  JIGs.append(create_jig_2(id=1, name="3FG", type=1, capacity=1, jig_offset=p[0,0,0,0,0,0]))
  JIGs.append(create_jig_2(id=2, name="jig input", type=2, capacity=1, jig_offset=p[0,0,0,0,0,-3.927]))
  JIGs.append(create_jig_2(id=3, name="jig output", type=3, capacity=1, jig_offset=p[0,0,0,0,0,0.78]))
  JIGs.append(create_jig_2(id=6, name="jig bin", type=6, capacity=1, jig_offset=p[0,0,0,0,0,0]))
  JIGs.append(create_jig_2(id=7, name="jig sarstedt racks", type=7, capacity=1, jig_offset=p[0,0,-0.02,0,0,0]))
  JIGs.append(create_jig_2(id=8, name="NoK Bin", type=8, capacity=1, jig_offset=p[0,0,0,0,0,0]))
  JIGs.append(create_jig_2(id=9, name="Pick bott jig", type=9, capacity=1, jig_offset=p[0,0,0,0,0,0]))
  JIGs.append(create_jig_2(id=10, name="Place bott jig", type=10, capacity=1, jig_offset=p[0,0,0,0,0,0]))
  JIGs.append(create_jig_2(id=11, name="bottle shake jig", type=11, capacity=1, jig_offset=p[0,0,0,0,0,0]))
  JIGs.append(create_jig_2(id=12, name="Pick Vial jig", type=12, capacity=1, jig_offset=p[0,0,0,0,0,0]))
  JIGs.append(create_jig_2(id=13, name="Place Vial jig", type=13, capacity=1, jig_offset=p[0,0,0,0,0,0]))
  JIGs.append(create_jig_2(id=14, name="Liquid transfer jig", type=14, capacity=1, jig_offset=p[0,0,0,0,0,0]))
  JIGs.append(create_jig_2(id=15, name="Pick station jig", type=15, capacity=1, jig_offset=p[0,0,0,0,0,0]))
  JIGs.append(create_jig_2(id=16, name="Place station jig", type=16, capacity=1, jig_offset=p[0,0,0,0,0,0]))
  JIGs.append(create_jig_2(id=17, name="Weigh station jig", type=17, capacity=1, jig_offset=p[0,0,0,0,0,0]))
  JIGs.append(create_jig_2(id=18, name="Pick station 1", type=18, capacity=1, jig_offset=p[0,0,0,0,0,0]))
  JIGs.append(create_jig_2(id=19, name="Pick station 2", type=19, capacity=1, jig_offset=p[0,0,0,0,0,0]))
  JIGs.append(create_jig_2(id=20, name="Pick station 3", type=20, capacity=1, jig_offset=p[0,0,0,0,0,0]))
  JIGs.append(create_jig_2(id=21, name="Tilt station jig", type=21, capacity=1, jig_offset=p[0,0,0,0,0,0]))
  $ 20 "Script: Powder_all_newspats.script"
  #global SERVER_IP   = "192.168.12.139"


  global tcp_dosing = p[0,0,0.15052,3.1415,0,0]
  global tcp_default = p[0,0,0.161,3.1415,0,0]

  global container_id = 0
  global powder_id  = 0
  global bulk_density = 0
  global H          = 0
  global H_c          = 0
  global mouth_d     = 0
  global mouth_sh    = 0
  global length_c     = 0
  global diameter   = 0
  global empty_weight_g  = 0
  global volume_ml    = 0
  global shape_code   = 0
  global flow_code   = 0
  global shape = ""
  global Flowability = ""
  global full_weight_g = 0
  global cent_edge = 0
  global pick_2_base = 0.2 # distance from tcp to base of picking table
  global wall_thickness = 0.002

  def read_db_data():

    socket_open(SERVER_IP, SERVER_PORT)
    sleep(0.5)
    socket_send_string("GET_DATACODE_FLOATS")
    sleep(5)

    local fl = socket_read_ascii_float(14)
    socket_close()

    global container_id = fl[1]
    global powder_id = fl[2]
    global bulk_density = fl[3]
    global H          = fl[4]/1000
    global H_c          = fl[5]/1000
    global mouth_d     = fl[6]/1000
    global mouth_sh    = fl[7]/1000
    global length_c     = fl[8]/1000
    global diameter   = fl[9]/1000
    global empty_weight_g = fl[10]
    global volume_ml    = fl[11]
    global full_weight_g = fl[12]
    global flow_code   = fl[13]
    global shape_code   = fl[14]

  	if (flow_code == 1.0):
  		global Flowability = "MEDIUM"
  	elif (flow_code == 2.0):
  		global Flowability = "LOW"
  	else:
  		global Flowability = "HIGH"
  	end

  	if ( shape_code == 1.0):
  		shape = "cylindrical"
  		cent_edge =  diameter
  	else:
  		shape = "cubical"
  		cent_edge =  length_c
  	end

  	read_spatula_data()

  end

  def send_picking_info(Pow_name, target_weight):
    socket_open(SERVER_IP, SERVER_PORT)
    cmd = "PICK:"+Pow_name+";"+to_str(target_weight)
    socket_send_string(cmd)
    sleep(0.1)
    socket_close()
  end

  #### POTS ####
  def tilt_send(angle):
  	socket_open(SERVER_IP, SERVER_PORT)
  	angle = 92.0 - angle
  	socket_send_string("TILT:"+to_str(angle))
  	sync()
  	sleep(0.5)
  	socket_close()
  end

  def CW_Rotate(angle):
  	socket_open(SERVER_IP, SERVER_PORT)
  	socket_send_string("CWROTATE:"+to_str(angle))
  	sync()
  	sleep(0.5)
  	socket_close()
  end

  def CCW_Rotate(angle):
  	socket_open(SERVER_IP, SERVER_PORT)
  	socket_send_string("CCWROTATE:"+to_str(angle))
  	sync()
  	sleep(0.5)
  	socket_close()
  end

  def CW_full_Rotate():
  	socket_open(SERVER_IP, SERVER_PORT)
  	socket_send_string("FULLROTATE:"+to_str(1))
  	sync()
  	sleep(0.5)
  	socket_close()
  end

  def CCW_full_Rotate():
  	socket_open(SERVER_IP, SERVER_PORT)
  	socket_send_string("FULLROTATE:"+to_str(-1))
  	sync()
  	sleep(0.5)
  	socket_close()
  end

  def tilt_to_home():
  	socket_open(SERVER_IP, SERVER_PORT)
  	socket_send_string("HOME")
  	sync()
  	sleep(0.5)
  	socket_close()
  end
  #######
  def vibration_1():
  	set_analog_out(0,0.4)
  	sleep(1)
  	set_analog_out(0,0.0)
  	sleep(0)
  end

  def vibration_2():
  	set_analog_out(0,0.4)
  	sleep(0.8)
  	set_analog_out(0,0.0)
  	sleep(0.2)
  end

  def vibration_3():
  	set_analog_out(0,0.4)
  	sleep(0.5)
  	set_analog_out(0,0.0)
  	sleep(0.3)
  end

  def vibration_4():
  	set_analog_out(0,0.4)
  	sleep(0.5)
  	set_analog_out(0, 0.0)
  	sleep(0.5)
  end

  def vibration_5():
  	set_analog_out(0,0.4)
  	sleep(0.2)
  	set_analog_out(0, 0.0)
  	sleep(0.8)
  end

  ##################

  global gear_2_holder = 0.018
  global hinge_2_base = 0.0421
  global TCP_2_tip_x = 0.0047
  global spatula_len = 0.182
  global spatula_offset = p[TCP_2_tip_x,0,spatula_len,0,0,0]
  global SPATULA_L_VOL_ML = 0.0
  global SPATULA_M_VOL_ML = 0.0
  global SPATULA_S_VOL_ML = 0.0
  global SPATULA_FLAT_M_VOL_ML  = 0.0
  global SPATULA_FLAT_S_VOL_ML  = 0.0

  global DB_SPATULA_L_DEPTH = 0.0
  global DB_SPATULA_M_DEPTH = 0.0
  global DB_SPATULA_S_DEPTH = 0.0
  global DB_SPATULA_FLAT_M_DEPTH = 0.0
  global DB_SPATULA_FLAT_S_DEPTH = 0.0
  global DB_SPATULA_L_MID = 0.0
  global DB_SPATULA_M_MID = 0.0
  global DB_SPATULA_S_MID = 0.0
  global DB_SPATULA_FLAT_M_MID = 0.0
  global DB_SPATULA_FLAT_S_MID = 0.0
  global DB_SPATULA_L_RY = 0.0
  global DB_SPATULA_M_RY = 0.0
  global DB_SPATULA_S_RY = 0.0
  global DB_SPATULA_FLAT_M_RY = 0.0
  global DB_SPATULA_FLAT_S_RY = 0.0

  def read_spatula_data():
  	socket_open(SERVER_IP, SERVER_PORT)
  	sleep(0.2)
  	socket_send_string("GET_SPATULA_FLOATS")
  	sleep(0.5)
  	local fl = socket_read_ascii_float(25)
  	socket_close()

  	global DB_SPATULA_L_DEPTH = fl[1]/1000
  	global DB_SPATULA_L_MID = fl[2]/2000
  	global SPATULA_L_VOL_ML = fl[3]
  	global DB_SPATULA_L_RY = fl[4]
  	global DB_SPATULA_M_DEPTH = fl[6]/1000
  	global DB_SPATULA_M_MID = fl[7]/2000
  	global SPATULA_M_VOL_ML = fl[8]
  	global DB_SPATULA_M_RY = fl[9]
  	global DB_SPATULA_S_DEPTH = fl[11]/1000
  	global DB_SPATULA_S_MID = fl[12]/2000
  	global SPATULA_S_VOL_ML = fl[13]
  	global DB_SPATULA_S_RY = fl[14]
  	global DB_SPATULA_FLAT_M_DEPTH = fl[16]/1000
  	global DB_SPATULA_FLAT_M_MID = fl[17]/2000
  	global SPATULA_FLAT_M_VOL_ML = fl[18]
  	global DB_SPATULA_FLAT_M_RY = fl[19]
  	global DB_SPATULA_FLAT_S_DEPTH = fl[21]/1000
  	global DB_SPATULA_FLAT_S_MID = fl[22]/2000
  	global SPATULA_FLAT_S_VOL_ML = fl[23]
  	global DB_SPATULA_FLAT_S_RY = fl[24]
  end

  def correction_reset():
  	global g_k = 0.0
  	global g_depth_corr = 0.0
  	global g_prev_cum_w = weight_value
  end

  def params_init():

  	global scoop_status= ""
  	global w_dosed_total = 0.0
  	global last_scale = 0.0
  	global tilt_angle_sent = 0.0
  	global level = 0.0
  	global target_g = 0.0
  	global angle_max = 65
  	global angle_min = 30
  	global gain_per_percent = (angle_max - angle_min)/100
  	global ry_deg_safe = 0
  	global ry_deg = 0
  	global delta_count=0

  	global scoop_ct = 0
  	global error_sum = 0.0
  	global error_sq_sum = 0.0
  	global scoop_g = 0.0

  	global g_k =0.0
  	global g_eta = 0.3

  	global g_gain_scale = 0.07
  	global g_k_min = 0.0
  	global g_k_max = 0.09

  	# ---------- Damping ----------
  	global g_alpha_under = 0.75   # aggressive when undershooting
  	global g_alpha_over  = 0.60   # conservative when overshooting

  	# ---------- Search ----------
  	global g_engagement_min = 0.05
  	global g_search_step = 0.01      # 3 mm

  	# ---------- Deadband ----------
  	global g_tol = 0.02               # 20 mg minimum
  	global g_tol_ratio = 0.05         # ±5% of target

  	# ---------- Limits ----------
  	global g_corr_max = 0.020         # 20 mm maximum correction

  	# ---------- States ----------
  	global g_depth_corr = 0.0
  	global g_prev_cum_w = -1.0
  	global z_ratio = 0.0
  	global z_offset = 0.0
  end

  def clamp(x, lo, hi):
  	if(x<lo):
  		return lo
  	elif (x>hi):
  		return hi
  	else:
  		return x
  	end
  end

  def compute_level_percent(W_now, weight_value):   # W_now = container+powder, weight_value = live scale reading
      global delta = weight_value - last_scale

      if (delta < 0.0):
          delta = 0.0
      end

      global w_dosed_total = w_dosed_total + delta
      global last_scale = weight_value     # update the last scale reading

      local W_eff = W_now - w_dosed_total
      if (W_eff <  empty_weight_g):
          W_eff =  empty_weight_g
      end

      # Compute powder level %
      level = 100.0 * (W_eff -  empty_weight_g) / (full_weight_g -  empty_weight_g)

      # Clamp to 0–100
      level = clamp(level, 0, 100)
    textmsg("deb 1 = ", level)
      return level
  end

  def deg2rad(d):
  	return d*3.141592/180
  end

  def my_abs(val):
  	if (val<0):
  		return -val
  	else:
  		return val
  	end
  end

  def compute_tilt_deg(level_percent):
  	angle = angle_min + gain_per_percent*(100.0-level_percent)

    	textmsg("deb 2 = ", angle)
  	return clamp(angle, angle_min, angle_max)
  end

  def tilt(level_percentage):
  	new_angle = compute_tilt_deg(level_percentage)
    	textmsg("deb angle 1 = ", new_angle)
  	global angle_rel = new_angle - tilt_angle_sent
    	textmsg("deb 2 = ", angle_rel)

  	if my_abs(angle_rel)>2.0:
    		textmsg("deb loop")
  		tilt_send(new_angle)
  		global angle_deg = new_angle
    		textmsg("deb 2 = ", angle_deg)
  		global tilt_angle_sent = new_angle
  		global p_center_vertical = center_pose()
  		global p_center = updated_center_pose(p_center_vertical, angle_deg)
  	end
    	textmsg("deb loop exit")

  	tilt_send(angle_deg)
    	textmsg("deb angle 2 =", angle_deg)

  end

  def compute_scoop_depth(level, weight_value, target_g):

      global scoop_depth_rel = ((100.0-level)/100.0)*(H-mouth_sh)

      if (g_prev_cum_w < 0):
          g_prev_cum_w = weight_value
          g_depth_corr = 0.0

      else:
          global scoop_g = weight_value - g_prev_cum_w
          g_prev_cum_w = weight_value

          local error = target_g - scoop_g
          local engagement = scoop_g / target_g

          local tol = g_tol_ratio * target_g
          if (tol < g_tol):
              tol = g_tol
          end
          if ((engagement < g_engagement_min) and (scoop_g < target_g)):
              g_depth_corr = g_depth_corr + g_search_step
          elif (my_abs(error) <= tol):
  			sync()
          else:
              local error_norm = my_abs(error / target_g)
              local g_target = clamp(g_gain_scale * error_norm,g_k_min,g_k_max)

              g_k = (1.0-g_eta) * g_k + g_eta * g_target
              if (error > 0):
                  local corr = g_k * error
                  g_depth_corr = g_depth_corr +g_alpha_under * corr
              else:
                  local corr = g_k * error
                  g_depth_corr = g_depth_corr +g_alpha_over * corr

              end
              g_depth_corr = clamp(g_depth_corr,-g_corr_max,g_corr_max)

          end
      end
      scoop_depth = scoop_depth_rel + g_depth_corr
      scoop_depth = clamp(scoop_depth, 0.0, H)
      return scoop_depth

  end

  def get_scoop_weight(spatula, bulk_density):

  	local vol = 0

  	if (spatula == "spatula_L"):
  		vol = SPATULA_L_VOL_ML
  		global spatula_depth = DB_SPATULA_L_DEPTH
  		global spatula_mid   = DB_SPATULA_L_MID
  		global spatula_ry    = DB_SPATULA_L_RY

  	elif (spatula == "spatula_M"):
  		vol = SPATULA_M_VOL_ML
  		global spatula_depth = DB_SPATULA_M_DEPTH
  		global spatula_mid   = DB_SPATULA_M_MID
  		global spatula_ry    = DB_SPATULA_M_RY

  	elif (spatula == "spatula_S"):
  		vol = SPATULA_S_VOL_ML
  		global spatula_depth = DB_SPATULA_S_DEPTH
  		global spatula_mid   = DB_SPATULA_S_MID
  		global spatula_ry    = DB_SPATULA_S_RY

  	elif (spatula == "spatula_flat_M"):
  		vol = SPATULA_FLAT_M_VOL_ML
  		global spatula_depth = DB_SPATULA_FLAT_M_DEPTH
  		global spatula_mid   = DB_SPATULA_FLAT_M_MID
  		global spatula_ry    = DB_SPATULA_FLAT_M_RY

  	elif (spatula == "spatula_flat_S"):
  		vol = SPATULA_FLAT_S_VOL_ML
  		global spatula_depth = DB_SPATULA_FLAT_S_DEPTH
  		global spatula_mid   = DB_SPATULA_FLAT_S_MID
  		global spatula_ry    = DB_SPATULA_FLAT_S_RY
  	else:
  		textmsg("Unknown spatula type")
  		return 0.0
  	end
  	global target_g = vol * bulk_density
  	return target_g

  end

  def select_spatula(Flowability, level, diff, bulk_density, mouth_d ):

      local k = 1.1
      global powder_height = (H  - mouth_sh ) * level/100

      if (Flowability == "LOW"):
          local gFM = get_scoop_weight("spatula_flat_M", bulk_density)
  		local mouth_ok_FM = (mouth_d >= 0.05)
  		local level_ok_FM = (spatula_mid  < powder_height)
          local diff_ok_FM  = (diff > k * gFM)
  		local flatM_ok = mouth_ok_FM and level_ok_FM and diff_ok_FM
          if (flatM_ok):
              return "spatula_flat_M"
          else:
              return "spatula_flat_S"
          end
      end

      local gL = get_scoop_weight("spatula_L", bulk_density)
      local mouth_ok_L = (mouth_d  >= 0.05)
      local level_ok_L = (spatula_mid < powder_height)
      local diff_ok_L  = (diff > k * gL)

      local large_ok = mouth_ok_L and level_ok_L and diff_ok_L
      local gM = get_scoop_weight("spatula_M", bulk_density)
      local level_ok_M = (spatula_mid < powder_height)
      local diff_ok_M  = (diff > k * gM)

      local medium_ok = level_ok_M and diff_ok_M

      if (large_ok):
          return "spatula_L"
      elif (medium_ok):
          return "spatula_M"
      else:
          return "spatula_S"
      end
  end

  def after_scoop():
  	set_tcp(tcp_dosing)
  	set_analog_out(0,0.0)
  	tilt_send(angle_deg)
  	sleep(0.5)
  	movel(lifted_pose, a=0.05, v=0.2)
  	movel(move_inside_spill, a=0.05, v=0.2)
  	set_analog_out(0,0.4)
  	if (Flowability == "LOW"):
  		movel(end_rel_tilted_level2, a=0.03, v=0.1)
  		sleep(0.5)
  		movel(move_inside_spill, a=0.05, v=0.2)
  	  	movel(pose_trans(move_inside_spill, p[0,0,0,0,0,2.0]), a=0.05, v=0.2)
  		#movel(tilted_pose_in_base2, a=0.05, v=0.2)
  	else:
  	    movel(pose_trans(move_inside_spill, p[0,0,0,0,0,2.0]), a=0.05, v=0.2)
  	    movel(move_inside_spill, a=0.05, v=0.2)
  	end
  	set_analog_out(0,0.0)
  	movel(lifted_pose, a=0.5, v=0.5)
  	tilt_to_home()
  	set_tcp(tcp_default)
  end

  def center_pose():
  	global p_translated = container_place
  	#global p_translated = pots_axis_temp

  	#cx = p_translated[0]
  	#cy = p_translated[1]
  	#cz = p_translated[2]

  	global p_center_vertical_temp = pose_trans(p_translated, p[0,0,0, deg2rad(90), 0, 0])
  	cx = p_center_vertical_temp[0]
  	cy = p_center_vertical_temp[1]
  	cz = p_center_vertical_temp[2]
  	rx = p_center_vertical_temp[3]
  	ry = p_center_vertical_temp[4]
  	rz = p_center_vertical_temp[5]

  	global p_center_vertical_temp = p[cx,cy,cz, 0, 0, rz]
  	trans_rel = p[0,0,-pick_2_base+H,0,0,0]
  	global p_center_vertical =  pose_trans(p_center_vertical_temp, trans_rel)
  	return p_center_vertical
  end

  def updated_center_pose(p_center_vertical, angle_deg):
  	hinge_pose = pose_trans(p_center_vertical, p[0,0,-hinge_2_base-gear_2_holder-H ,0,0,0])
  	local_rel = pose_trans(pose_inv(hinge_pose), p_center_vertical)

  	rot_tilt = p[0,0,0, -deg2rad(angle_deg),0,0]
  	local_rel_tilted = pose_trans(rot_tilt, local_rel)

  	global p_center = pose_trans(hinge_pose, local_rel_tilted)
  	return p_center
  end

  def scoop_powder(p_center):
  	vibration_voltage = 0.4
  	global scoop_radius_default = 0.0

  	scoop_radius_default = mouth_d /2 - spatula_depth - wall_thickness
  	scoop_safe_entry_pose = pose_trans(p_center, p[-TCP_2_tip_x,0,spatula_len+0.05,0,0,0])
  	scoop_entry_pose = pose_trans(p_center, p[-TCP_2_tip_x,0,spatula_len,0,0,0])

  	movel(scoop_safe_entry_pose, a=0.1, v=0.25)
  	movel(scoop_entry_pose, a=0.1, v=0.25)

  	scoop_start_rel_int = p[0, 0, -mouth_sh , 0, 0, 0]
  	scoop_start_pose_int = pose_trans(scoop_entry_pose, scoop_start_rel_int)


  	#local ry_deg = map_tilt_to_ry_deg(angle_deg,level)
  	#local ry_result = map_tilt_to_ry_deg(angle_deg,level)

  	#global scoop_depth = compute_scoop_depth(level,weight_value, target_g)

  	global ry = deg2rad(90-angle_deg)

  	#global ry_safe = ry_result[0]
  	#global ry = deg2rad(ry_result[1])

  	if (spatula_mid < powder_height):

  		global total_depth = mouth_sh + scoop_depth + spatula_mid
  		global total_depth = clamp(total_depth, 0, H - spatula_mid)

  		safe_scoop_pivot = (mouth_d  - spatula_depth-wall_thickness)/(total_depth)
  		global ry_safe = asin(safe_scoop_pivot)

  		scoop_start_rel = p[scoop_radius_default, 0, -total_depth, 0, 0, 0]

  		rot_mid = p[0, 0, 0, 0, 0, 0.785]
  		rot_end = p[0, 0, 0, 0, 0, 1.5708]

  		scoop_via_rel = pose_trans(rot_mid, scoop_start_rel)
  		scoop_end_rel = pose_trans(rot_end, scoop_start_rel)

  		scoop_start_pose = pose_trans(scoop_entry_pose, scoop_start_rel)
  		scoop_via_pose = pose_trans(scoop_entry_pose, scoop_via_rel)
  		scoop_end_pose = pose_trans(scoop_entry_pose, scoop_end_rel)


  			if (Flowability == "LOW" and level <= 50):
  				movel(pose_trans(scoop_start_pose_int,p[0,0,0,0,0,-1.5708]), a=0.1, v=0.25)
  				local spatula_base = pose_trans(scoop_entry_pose, p[0, 0, -H+wall_thickness, 0, 0, 0])
  				local scrape_pivot = pose_trans(scoop_entry_pose, p[0,0, -spatula_len,0,0,0])

  				global sticky_in_angle = -atan((cent_edge/2-spatula_depth)/H)
  				spatula_tilt_rel = pose_trans(pose_inv(scrape_pivot), spatula_base)

  				spatula_tilt = pose_trans(spatula_tilt_rel, p[0, 0, 0, 0, sticky_in_angle, 0])
  				global tilted_pose = pose_trans(scrape_pivot, p[0,0,0,spatula_tilt[3],spatula_tilt[4], spatula_tilt[5]])

  				global tilted_pose = pose_trans(tilted_pose, p[0,0,spatula_len-H+wall_thickness,0,0,0])
  				global rotate_90=pose_trans(tilted_pose,p[0,0,0,0,0,-1.5708])
  				movel(rotate_90,a=0.1, v=0.25)
  				CW_full_Rotate()
  				movel(scoop_start_pose, a=0.1, v=0.25)
  			else:
  				movel(scoop_start_pose_int, a=0.1, v=0.25)
  				movel(scoop_start_pose, a=0.1, v=0.25)
  				CW_full_Rotate()
  			end

  		movec(scoop_via_pose, scoop_end_pose, a=0.05, v=0.04)
  		#sleep(1.0)

  		# safe_retention
  		local pivot_pose = pose_trans(scoop_end_pose, p[0,0,total_depth-spatula_len,0,0,0])
  		local end_rel = pose_trans(pose_inv(pivot_pose), scoop_end_pose)
  		local end_rel_tilted = pose_trans(end_rel, p[0, 0, 0, 0, ry_safe-deg2rad(spatula_ry), 0])
  		local tilted_pose_in_base = pose_trans(pivot_pose, p[0,0,0,end_rel_tilted[3],end_rel_tilted[4], end_rel_tilted[5]])
  		local tilted_pose_in_base = pose_trans(tilted_pose_in_base, p[0, 0, spatula_len-total_depth, 0, 0, 0])
  		# sptula pivoted around the container rim of the mouth at ry_safe
  		movel(tilted_pose_in_base, a=0.03, v=0.1)

  		global safe_x = sin(ry_safe)*(total_depth-mouth_sh - (mouth_d - spatula_depth)*tan(ry_safe/2))
  		global safe_z = cos(ry_safe)*(total_depth-mouth_sh - (mouth_d - spatula_depth)*tan(ry_safe/2))

  		local safe_up = pose_trans(tilted_pose_in_base, p[-safe_x,0,safe_z,0,0,0])
  		movel(safe_up, a=0.03, v=0.1)

  		# full exit
  		local pivot_pose2 = pose_trans(scoop_entry_pose, p[0,0,-spatula_len,0,0,0])
  		local end_rel2 = pose_trans(pose_inv(pivot_pose2), tilted_pose_in_base)
  		#popup("is the spatula crashing front? ", blocking = True)
  		local end_rel_tilted2 = pose_trans(end_rel2, p[0, 0, 0, 0, ry-ry_safe-deg2rad(spatula_ry), 0])

  	else : # emptying logic
  		#CCW_full_Rotate()

  		spatula_base = pose_trans(scoop_entry_pose, p[0, 0, -H+wall_thickness, 0, 0, 0])
  		local pivot_pose2 = pose_trans(scoop_entry_pose, p[0,0,-spatula_len,0,0,0])
  		# tilt inwards
  		global in_angle = -atan((cent_edge/2-spatula_depth)/H)
  		spatula_tilt_rel = pose_trans(pose_inv(pivot_pose2), spatula_base)

  		spatula_tilt = pose_trans(spatula_tilt_rel, p[0, 0, 0, -in_angle, 0, 0])
  		global tilted_pose = pose_trans(pivot_pose2, p[0,0,0,spatula_tilt[3],spatula_tilt[4], spatula_tilt[5]])

  		global tilted_pose = pose_trans(tilted_pose, p[0,0,spatula_len-H+wall_thickness,0,0,0])

  		movel(tilted_pose,a=0.1, v=0.25)
  		CW_full_Rotate()
  		sleep(1)
  		rotate90=pose_trans(tilted_pose,p[0,0,0,0,0,1.5708])

  		#sleep(1)
  		#Rotate()
  		#sleep(0.2)
  		movel(rotate90, a=0.1, v=0.1)
  		#popup("is the spatula crashing front? ", blocking = True)
  		movel(pose_trans(scoop_start_pose_int,p[0,0,0,0,0,1.5708]), a=0.03, v=0.1)
  		# full exit
  		#local pivot_pose2 = pose_trans(scoop_entry_pose, p[0,0,-spatula_len,0,0,0])
  		local end_rel2 = pose_trans(pose_inv(scoop_entry_pose), rotate90)
  		local end_rel_tilted2 = pose_trans(end_rel2, p[0, 0, 0, 0, ry-in_angle-deg2rad(spatula_ry), 0])
  	end

  	# exit flat spoon
  	global tilted_pose_in_base2 = pose_trans(pivot_pose2, p[0,0,0,end_rel_tilted2[3],end_rel_tilted2[4], end_rel_tilted2[5]])
  	global tilted_pose_in_base2 = pose_trans(tilted_pose_in_base2, p[0, 0, spatula_len-spatula_mid, 0, 0, 0])
  	# spaula exited at center of the mouth at ry
  	movel(tilted_pose_in_base2, a=0.03, v=0.1)

  	if(spatula == "spatula_S"):
  		if(level>=80):
  			global z_ratio = 0.0
  		elif(level == 0.0):
  			global z_ratio = 1.0
  		else:
  			global z_ratio = (80-level)/80
  		end
  		z_offset = 4*spatula_mid*z_ratio
  	elif(spatula == "spatula_flat_S"):
  		if(level>=50):
  			global z_ratio = 0.0
  		elif(level == 0.0):
  			global z_ratio = 1.0
  		else:
  			global z_ratio = (50-level)/50
  		end
  		z_offset = 4*spatula_mid*z_ratio
  	else:
  	    z_offset = 0.0
  	end

  	global move_inside_spill = pose_trans(tilted_pose_in_base2, p[0,0,-z_offset,0,0,0])
  	movel(move_inside_spill, a=0.03, v=0.1)

  	if(scoop_status== "normal"):
  		vib_thread=True
  		if (spatula=="spatula_S"):
  			vibration_3()
  			local ry_level = deg2rad(5)
  		elif(spatula=="spatula_flat_S" or spatula=="spatula_flat_M"):
  			vibration_3()
  			local ry_level = deg2rad(5)
  		else:
  			set_analog_out(0,0.4)
  			local ry_level = deg2rad(15)
  		end

  		# remove excess
  		local pivot_pose_level = pose_trans(move_inside_spill, p[0,0,-spatula_len,0,0,0])
  		local end_rel_level = pose_trans(pose_inv(pivot_pose_level), move_inside_spill)
  		local end_rel_tilted_level = pose_trans(end_rel_level, p[0, 0, 0, 0, -ry_level, 0])
  		global end_rel_tilted_level2 = pose_trans(pivot_pose_level, p[0, 0, 0,end_rel_tilted_level[3],end_rel_tilted_level[4], end_rel_tilted_level[5]])
  		global end_rel_tilted_level2 = pose_trans(end_rel_tilted_level2, p[0,0,spatula_len,0,0,0])
  		movel(end_rel_tilted_level2, a=0.03, v=0.1)

  		if (spatula == "spatula_flat_S" or spatula == "spatula_flat_M"):
  			vib_thread=False
  			set_analog_out(0, 0.0)
  		end
  	else:
  		set_analog_out(0, 0.0)
  	end
  	movel(tilted_pose_in_base2, a=0.03, v=0.1)
  	set_analog_out(0, 0.0)
  	vib_thread=False
  	global lifted_pose = pose_trans(tilted_pose_in_base2, p[-0.04,0,0.04,0,0,0]) # safety distance away from the container

  	movel(lifted_pose, a=0.03, v=0.1)
  	tilt_to_home()
  end

  def auto_tilt_and_scoop(W_now, target_weight, weight_value):
  	set_tcp(tcp_dosing)
  	#global level = compute_level_percent(W_now, weight_value)

  	global spatula = select_spatula(Flowability, level, diff, bulk_density, mouth_d )
  	textmsg("deb 4 = ", spatula)
  	global target_g = get_scoop_weight(spatula, bulk_density)
  	textmsg("deb 5 = ", target_g)

  	global scoop_depth = compute_scoop_depth(level, weight_value, target_g)
    	textmsg("deb 6 = ", scoop_depth)
  	tilt(level)

  	scoop_powder(p_center)

  	#textmsg("deb 7 - sucess")
   	set_tcp(tcp_default)
  end
  $ 21 "Script: Weight_scale_socket_s.script"
  global s_depth = 0
  global s_length =0
  global s_volume = 0
  global ry_theta  = 0

  def get_weight():
  	socket_open(SERVER_IP,SERVER_PORT)
  	#sleep(0.2)
  	textmsg("socket opened successfully!")
  	socket_send_string("GET_WEIGHT")
  	#sleep(0.2)
  	sync()
  	receiveFromServ = socket_read_ascii_float(1)
  	#sleep(1)
  	while (receiveFromServ[0] < 1):
  		receiveFromServ = socket_read_ascii_float(1)
  		sleep(0.01)
  	end
  	textmsg("Received weight:", receiveFromServ[1])
  	#sleep(0.2)
  	socket_close()
  	#sleep(0.2)
  	return receiveFromServ[1]
  end

  def tare_scale():
  	socket_open(SERVER_IP,SERVER_PORT)
  	socket_send_string("TARE")
  	sleep(2)
  	socket_close()
  end

  def zero_scale():
  	socket_open(SERVER_IP,SERVER_PORT)
  	socket_send_string("ZERO")
  	sleep(0.5)
  	socket_close()
  end

  def log_weight():
  	socket_open(SERVER_IP,SERVER_PORT)
  	socket_send_string("LOG_WEIGHT")
  	sleep(0.5)
  	socket_close()
  end

  def send_target_info():
  	socket_open(SERVER_IP,SERVER_PORT)
  	socket_send_string("SET_TARGET:" + to_str(target_weight))
  	sleep(0.2)
  	socket_close()
  end
  def send_powder_info():
  	socket_open(SERVER_IP,SERVER_PORT)
  	socket_send_string("SET_POWDER:" + Pow_name)
  	sleep(0.2)
  	socket_close()
  end
  def send_spatula_info():
  	socket_open(SERVER_IP,SERVER_PORT)
  	socket_send_string("SET_SPATULA:" + spatula)
  	#sleep(1)

  	#local fl = socket_read_ascii_float(4)

    	#global s_depth = fl[1]
    	#global s_length = fl[2]
   	#global s_volume = fl[3]
   	#global ry_theta  = fl[4]
  	sleep(0.2)
  	socket_close()
  end

  def send_level_info():
  	socket_open(SERVER_IP,SERVER_PORT)
  	socket_send_string("SET_LEVEL:" + to_str(level))
  	sleep(0.2)
  	socket_close()
  end

  def get_cont_weight():
    socket_open(SERVER_IP, SERVER_PORT)
    #rq_open_and_wait()
    cmd = "GET_CONT_WEIGHT"
    socket_send_string(cmd)
    sync()
    sleep(0.5)
    receiveFromSer = socket_read_ascii_float(1)
    socket_close()
    return receiveFromSer[1]
  end

  $ 22 "Script: swab_sampling.script"
  def connect2server():
  	IP="192.168.12.139"
  	port=3002
  	cntd=False
  	while(cntd==False):
  		cntd=socket_open(IP,port,"PYSERV")
  		textmsg("Connected to server")
  	end
  	socket_send_string("SCAN_TARGET","PYSERV")
  	#sleep(200)
  	#resp=socket_read_binary_integer(1,"PYSERV",timeout=-1)
  	#textmsg("Response",resp)
  	#if(resp[0]==1):
  		#motion=True
  		#while(motion == True):
  			#msg=socket_read_ascii_float(6,"PYSERV",timeout=-1)
  			#textmsg("msg recieved",msg)
  			#if(msg[0]==6):
   	    		#	textmsg("INSIDE MOVE")
  	    		#	trg_pose=p[msg[1],msg[2],msg[3],msg[4],msg[5],msg[6]]
  	    		#	movel(trg_pose,a=0.2,v=0.25)
  			#	socket_send_string("ACKNO","PYSERV")
  	  		#else:
  				motion=False
  			#end
  		#end
  	#	resp=""
  	textmsg("Python taking over")
  	finish_msg=socket_read_string("PYSERV",timeout=-1)
  	textmsg("Motion Finished msg: ", finish_msg)

  	#end
  	textmsg("Motion Finished")
  	socket_close()
  end
  $ 23 "BeforeStarts"
  $ 24 "uLM"
  $ 25 "CMD_Stop≔ False "
  global CMD_Stop=  False
  $ 26 "CMD_Abort≔ False "
  global CMD_Abort=  False
  $ 27 "CMD_Clear≔ False "
  global CMD_Clear=  False
  $ 28 "STATE≔1"
  global STATE=1
  $ 29 "STATE_Info≔''"
  global STATE_Info=""
  $ 30 "ARM_Referenced≔ False "
  global ARM_Referenced=  False
  $ 31 "zero_ftsensor()"
  zero_ftsensor()
  $ 32 "poses init"
  $ 33 "PSE_A≔p[0,0,0,0,0,0]"
  global PSE_A=p[0,0,0,0,0,0]
  $ 34 "PSE_A_H≔p[0,0,0,0,0,0]"
  global PSE_A_H=p[0,0,0,0,0,0]
  $ 35 "PSE_R≔p[0,0,0,0,0,0]"
  global PSE_R=p[0,0,0,0,0,0]
  $ 36 "PSE_R_H≔p[0,0,0,0,0,0]"
  global PSE_R_H=p[0,0,0,0,0,0]
  $ 37 "PSE_T≔p[0,0,0,0,0,0]"
  global PSE_T=p[0,0,0,0,0,0]
  $ 38 "PSE_T_H≔p[0,0,0,0,0,0]"
  global PSE_T_H=p[0,0,0,0,0,0]
  $ 39 "PSE_C_E≔p[0,0,0,0,0,0]"
  global PSE_C_E=p[0,0,0,0,0,0]
  $ 40 "PSE_C_H≔p[0,0,0,0,0,0]"
  global PSE_C_H=p[0,0,0,0,0,0]
  $ 41 "PSE_C_S≔p[0,0,0,0,0,0]"
  global PSE_C_S=p[0,0,0,0,0,0]
  $ 42 "init_home_by_cartesian_pose(p[0,-0.400,0.300,0,0,0])"
  init_home_by_cartesian_pose(p[0,-0.400,0.300,0,0,0])
  $ 43 "Clearing"
  $ 44 "reset_error()"
  reset_error()
  $ 45 "reset_warning()"
  reset_warning()
  $ 46 "uGo"
  $ 48 "ugo_init( True ,'http://192.168.12.120:10001')"
  ugo_init(  True  ,"http://192.168.12.120:10001")
  $ 49 "ugo_update_outputs()"
  ugo_update_outputs()
  $ 50 "App"
  $ 51 "'ADD APPLICATION SPECIFIC COMMANDS'"
  # 'ADD APPLICATION SPECIFIC COMMANDS'
  $ 52 "Tools"
  $ 53 "OBJ_Picked≔gripper_has_object()"
  global OBJ_Picked=gripper_has_object()
  $ 54 "If OBJ_Picked"
  if (OBJ_Picked):
    # begin: URCap Program Node
    #   Source: Robotiq_Grippers, 3.17.0.105337, Robotiq Inc.
    #   Type: Gripper Activate
    $ 55 "Gripper Activate"

    kill rq_gripper_communication_thread
    rq_gripper_communication_thread_started = False
    rq_close_gripper_socket("1")
    rq_close_gripper_socket("2")
    rq_close_gripper_socket("3")
    rq_close_gripper_socket("4")

    rq_init_comm_if_connected(9, "1")
    rq_init_comm_if_connected(2, "2")
    rq_init_comm_if_connected(3, "3")
    rq_init_comm_if_connected(4, "4")
    rq_print_connected_grippers()
    rq_gripper_communication_thread = run rq_gripper_communication()

    while(not rq_gripper_communication_thread_started):
        sleep(0.008)
    end

    rq_set_max_current_for_all_grippers()

    reset_and_activate = False

    rq_activate_all_grippers(False)
    # end: URCap Program Node
  else:
    $ 56 "Else" "noBreak"
    # begin: URCap Program Node
    #   Source: Robotiq_Grippers, 3.17.0.105337, Robotiq Inc.
    #   Type: Gripper Activate
    $ 57 "Gripper Reset and Activate"

    kill rq_gripper_communication_thread
    rq_gripper_communication_thread_started = False
    rq_close_gripper_socket("1")
    rq_close_gripper_socket("2")
    rq_close_gripper_socket("3")
    rq_close_gripper_socket("4")

    rq_init_comm_if_connected(9, "1")
    rq_init_comm_if_connected(2, "2")
    rq_init_comm_if_connected(3, "3")
    rq_init_comm_if_connected(4, "4")
    rq_print_connected_grippers()
    rq_gripper_communication_thread = run rq_gripper_communication()

    while(not rq_gripper_communication_thread_started):
        sleep(0.008)
    end

    rq_set_max_current_for_all_grippers()

    reset_and_activate = True

    rq_activate_all_grippers(True)
    # end: URCap Program Node
  end
  $ 58 "zero_ftsensor()"
  zero_ftsensor()
  $ 59 "EXTT"
  $ 60 "Set GRP_3F_Enable=Off"
  set_standard_digital_out(4, False)
  $ 61 "Set BarcodeTrigger=Off"
  set_standard_digital_out(6, False)
  $ 62 "Set GRP_3F_Decap=Off"
  set_standard_digital_out(3, False)
  $ 63 "Set GRP_3F_Cap=Off"
  set_standard_digital_out(2, False)
  $ 64 "Set GRP_3F_Open=Off"
  set_standard_digital_out(5, False)
  $ 65 "PSE_T≔get_tool_free_pose(dir=[0,0,0.150], move_in_base_frame=True)"
  global PSE_T=get_tool_free_pose(dir=[0,0,0.150], move_in_base_frame=True)
  $ 66 "If is_reachable(Base_const, [PSE_T])"
  if (is_reachable(p[0.0,0.0,0.0,0.0,0.0,0.0], [PSE_T])):
    $ 67 "MoveL"
    $ 68 "PSE_T" "breakAfter"
    movel(PSE_T, a=1.2, v=0.15)
  end
  $ 69 "powder dispensing variable init"
  $ 70 "Start_thread≔ False "
  global Start_thread=  False
  $ 71 "vib_thread≔ False "
  global vib_thread=  False
  $ 72 "w_full_thread≔ False "
  global w_full_thread=  False
  $ 73 "Picking≔ False "
  global Picking=  False
  $ 74 "d_cc≔0.07"
  global d_cc=0.07
  $ 75 "kp≔0.0035"
  global kp=0.0035
  $ 76 "ki≔0.0001"
  global ki=0.0001
  $ 77 "kd≔0.003"
  global kd=0.003
  $ 78 "dt≔0.2"
  global dt=0.2
  $ 79 "Integral_error≔0"
  global Integral_error=0
  $ 80 "current_error≔0"
  global current_error=0
  $ 81 "previous_error≔0"
  global previous_error=0
  $ 82 "tilt_increment≔0"
  global tilt_increment=0
  $ 83 "tilt_angle≔0"
  global tilt_angle=0
  $ 84 "diff≔0"
  global diff=0
  $ 85 "tilt_to_home()"
  tilt_to_home()
  $ 86 "params_init()"
  params_init()
  $ 87 "switch_spat_M≔ True "
  global switch_spat_M=  True
  $ 88 "switch_spat_S≔ True "
  global switch_spat_S=  True
  $ 89 "switch_spat_F_M≔ True "
  global switch_spat_F_M=  True
  $ 90 "switch_spat_F_S≔ True "
  global switch_spat_F_S=  True
  $ 91 "last_scale≔0"
  global last_scale=0
  $ 858 "Thread_1"
  thread Thread_1():
    while (True):
      $ 859 "Dosing Weight"
      $ 860 "If Start_thread≟ True "
      if (Start_thread ==   True  ):
        $ 861 "weight_value≔get_weight()"
        global weight_value=get_weight()
        $ 862 "diff≔target_weight-weight_value"
        global diff=target_weight-weight_value
        $ 863 "Wait: 0.2"
        sleep(0.2)
        $ 864 "sync()"
        sync()
      end
      $ 865 "sync()"
      sync()
    end
  end
  threadId_Thread_1 = run Thread_1()
  $ 866 "Thread_2"
  thread Thread_2():
    while (True):
      $ 867 "Vibration motor"
      $ 868 "Loop vib_thread≟ True "
      thread Thread_while_868():
        while (True):
          $ 869 "diff≔target_weight-weight_value"
          global diff=target_weight-weight_value
          $ 870 "If diff>0.02 and spatula≠'spatula_flat_S' "
          global thread_flag_870=0
          thread Thread_if_870():
            $ 872 "Set AO[0]=4.0"
            set_standard_analog_out(0, 0.4)
            thread_flag_870 = 1
          end
          if (diff>0.02  and  spatula != "spatula_flat_S" ):
            global thread_handler_870=run Thread_if_870()
            while (thread_flag_870 == 0):
              if not(diff>0.02  and  spatula != "spatula_flat_S" ):
                kill thread_handler_870
                thread_flag_870 = 2
              else:
                sync()
              end
            end
          else:
            thread_flag_870 = 2
          end
          if (thread_flag_870 == 2):
            $ 873 "ElseIf diff>0.02 and spatula≟'spatula_flat_S'"
            if (diff>0.02 and spatula == "spatula_flat_S"):
              $ 874 "vibration_3()"
              vibration_3()
            else:
              $ 875 "ElseIf diff≤0.03"
              global thread_flag_875=0
              thread Thread_if_875():
                $ 876 "vibration_2()"
                vibration_2()
                thread_flag_875 = 1
              end
              if (diff <= 0.03):
                global thread_handler_875=run Thread_if_875()
                while (thread_flag_875 == 0):
                  if not(diff <= 0.03):
                    kill thread_handler_875
                    thread_flag_875 = 2
                  else:
                    sync()
                  end
                end
              else:
                thread_flag_875 = 2
              end
              if (thread_flag_875 == 2):
                $ 877 "Else" "noBreak"
                $ 878 "Set AO[0]=0.0"
                set_standard_analog_out(0, 0.0)
              end
            end
          end
        end
      end
      if (vib_thread ==   True  ):
        global thread_handler_868=run Thread_while_868()
        while (vib_thread ==   True  ):
          sync()
        end
        kill thread_handler_868
      end
      $ 879 "sync()"
      sync()
    end
  end
  threadId_Thread_2 = run Thread_2()
  $ 880 "Thread_3"
  thread Thread_3():
    while (True):
      $ 881 "Container weight"
      $ 882 "If w_full_thread≟ True "
      if (w_full_thread ==   True  ):
        $ 883 "aa_weight_cont≔get_cont_weight()"
        global aa_weight_cont=get_cont_weight()
        $ 884 "Wait: 0.2"
        sleep(0.2)
        $ 885 "sync()"
        sync()
      end
      $ 886 "sync()"
      sync()
    end
  end
  threadId_Thread_3 = run Thread_3()
  while (True):
    $ 92 "Robot Program"
    $ 93 "MAIN"
    $ 94 "command_manager(external_control='uGO', cond_suspend=(ITM_Manipulated and AMR_AtTarget and AMR_Charging and AMR_Battery<40), cond_unsuspend=(AMR_Battery≟60))"
    command_manager(external_control="uGO", cond_suspend=(ITM_Manipulated  and  AMR_AtTarget  and  AMR_Charging  and  AMR_Battery<40), cond_unsuspend=(AMR_Battery == 60))
    $ 95 "log_state(STATE_Info)"
    log_state(STATE_Info)
    $ 96 "Switch STATE"
    switch_1 = STATE
    $ 97 "Case 1"
    if (1 == switch_1):
      $ 98 "Stopping"
      $ 99 "STATE_Info≔'Stopping'"
      global STATE_Info="Stopping"
      $ 100 "end_freedrive_mode()"
      end_freedrive_mode()
      $ 101 "Set"
      set_tcp(p[0.0,0.0,0.161,3.1415,0.0,0.0])
      $ 102 "PSE_T≔get_tool_free_pose(dir=[0,0,0.150], move_in_base_frame=True)"
      global PSE_T=get_tool_free_pose(dir=[0,0,0.150], move_in_base_frame=True)
      $ 103 "If is_reachable(Base_const, [PSE_T])"
      if (is_reachable(p[0.0,0.0,0.0,0.0,0.0,0.0], [PSE_T])):
        $ 104 "MoveL"
        $ 105 "PSE_T" "breakAfter"
        movel(PSE_T, a=1.2, v=0.15)
      end
      $ 106 "do_transition(keep_rxry=OBJ_Picked, r=0)"
      do_transition(keep_rxry=OBJ_Picked, r=0)
      $ 115 "Call Sub_AMR_MiR_V3"
      Sub_AMR_MiR_V3()
      $ 116 "If stopping() and AMR_Done"
      if (stopping()  and  AMR_Done):
        $ 117 "STATE≔2"
        global STATE=2
        $ 118 "ugo_update_outputs()"
        ugo_update_outputs()
      end
    elif (2 == switch_1):
      $ 119 "Case 2"
      $ 120 "Stopped"
      $ 121 "STATE_Info≔'Stopped'"
      global STATE_Info="Stopped"
      $ 122 "Call Sub_AMR_MiR_V3"
      Sub_AMR_MiR_V3()
      $ 123 "If CMD_Reset  or PB_Start"
      if (CMD_Reset   or  get_standard_digital_in(0)):
        $ 124 "STATE≔3"
        global STATE=3
        $ 125 "ugo_update_outputs()"
        ugo_update_outputs()
      end
    elif (3 == switch_1):
      $ 126 "Case 3"
      $ 127 " Resetting"
      $ 128 "STATE_Info≔'Resetting'"
      global STATE_Info="Resetting"
      $ 129 "uML"
      $ 130 "reset_error()"
      reset_error()
      $ 131 "reset_warning()"
      reset_warning()
      $ 132 "PROCESS_Step≔0"
      global PROCESS_Step=0
      $ 133 "PROCESS_Info≔''"
      global PROCESS_Info=""
      $ 134 "ARM_Referenced≔ False "
      global ARM_Referenced=  False
      $ 135 "WRK_Done≔ False "
      global WRK_Done=  False
      $ 136 "ITM_Prepared≔ False "
      global ITM_Prepared=  False
      $ 137 "ITM_Manipulated≔ False "
      global ITM_Manipulated=  False
      $ 138 "STP≔0"
      global STP=0
      $ 139 "Action≔0"
      global Action=0
      $ 140 "Action_Info≔''"
      global Action_Info=""
      $ 141 "ITM_ID≔0"
      global ITM_ID=0
      $ 142 "JIG≔0"
      global JIG=0
      $ 143 "JIG_Slot≔0"
      global JIG_Slot=0
      $ 144 "Task_info≔''"
      global Task_info=""
      $ 145 "Set"
      set_tcp(p[0.0,0.0,0.161,3.1415,0.0,0.0])
      $ 146 "App"
      $ 147 "'ADD APPLICATION SPECIFIC COMMANDS'"
      # 'ADD APPLICATION SPECIFIC COMMANDS'
      $ 148 "OBJ_Type≔0"
      global OBJ_Type=0
      $ 149 "OBJ_Nbr≔0"
      global OBJ_Nbr=0
      $ 150 "If CNT_Rack_Output≥50"
      if (CNT_Rack_Output >= 50):
        $ 151 "CNT_Rack_Output≔0"
        global CNT_Rack_Output=0
      end
      $ 152 "TASK≔struct(ID=0, NAVI=struct(target=0, footprint=0, protectiveOff=0, dock=0), WORK=struct(ITM_ID_Src=0, JIG_ID_Src=0, OBJ_Nbr_Src=0, ACT_Src=0, ITM_ID_Tgt=0, JIG_ID_Tgt=0, OBJ_Nbr_Tgt=0, ACT_Tgt=0, OBJ_Type=0))"
      global TASK=struct(ID=0, NAVI=struct(target=0, footprint=0, protectiveOff=0, dock=0), WORK=struct(ITM_ID_Src=0, JIG_ID_Src=0, OBJ_Nbr_Src=0, ACT_Src=0, ITM_ID_Tgt=0, JIG_ID_Tgt=0, OBJ_Nbr_Tgt=0, ACT_Tgt=0, OBJ_Type=0))
      $ 153 "Call Sub_AMR_MiR_V3"
      Sub_AMR_MiR_V3()
      $ 154 "If resetting() and AMR_Done"
      if (resetting()  and  AMR_Done):
        $ 155 "STATE≔4"
        global STATE=4
        $ 156 "ugo_update_outputs()"
        ugo_update_outputs()
      end
    elif (4 == switch_1):
      $ 157 "Case 4"
      $ 158 "Idle"
      $ 159 "STATE_Info≔'Idle'"
      global STATE_Info="Idle"
      $ 160 "If CMD_Start"
      if (CMD_Start):
        $ 161 "STATE≔5"
        global STATE=5
        $ 162 "ugo_update_outputs()"
        ugo_update_outputs()
      end
    elif (5 == switch_1):
      $ 163 "Case 5"
      $ 164 "Starting"
      $ 165 "STATE_Info≔'Starting'"
      global STATE_Info="Starting"
      $ 166 "'ADD COMMANDS WHAT TO START WITH'"
      # 'ADD COMMANDS WHAT TO START WITH'
      $ 167 "Call Sub_AMR_MiR_V3"
      Sub_AMR_MiR_V3()
      $ 168 "get ugo data"
      $ 169 "Assign Tasks"
      $ 170 "TASK.ID = ugo_get_task()"
      TASK.ID = ugo_get_task()
      $ 171 "If TASK.ID≟1"
      if (TASK.ID == 1):
        $ 172 "Task_info≔'Charge'"
        global Task_info="Charge"
        $ 173 "Parameters"
        $ 174 "AMR_PosTarget≔1"
        global AMR_PosTarget=1
      else:
        $ 175 "ElseIf TASK.ID≟9"
        if (TASK.ID == 9):
          $ 176 "'Pick Sarstedt Rack from Variable source'"
          # 'Pick Sarstedt Rack from Variable source'
          $ 177 "Task_info≔'Navigate to Target'"
          global Task_info="Navigate to Target"
          $ 178 "Parameters"
          $ 179 "AMR_PosTarget≔UGO.read_input('00','ITM_ID')"
          global AMR_PosTarget=UGO.read_input("00","ITM_ID")
        else:
          $ 180 "ElseIf TASK.ID≟13"
          if (TASK.ID == 13):
            $ 181 "Task_info≔'Dose Powder'"
            global Task_info="Dose Powder"
            $ 182 "Parameters"
            $ 183 "ITM_ID≔1"
            global ITM_ID=1
            $ 184 "W_now≔(UGO.read_input('00','Container_weight'))/1000"
            global W_now=(UGO.read_input("00","Container_weight"))/1000
            $ 185 "Pow_name≔(UGO.read_input('00','Powder_name'))"
            global Pow_name=(UGO.read_input("00","Powder_name"))
            $ 186 "target_weight≔(UGO.read_input('00','Target_weight'))/1000"
            global target_weight=(UGO.read_input("00","Target_weight"))/1000
            $ 187 "params_init()"
            params_init()
            $ 188 "send_picking_info(Pow_name,target_weight)"
            send_picking_info(Pow_name,target_weight)
            $ 190 "OBJ_Type≔6"
            global OBJ_Type=6
            $ 191 "JIG≔17"
            global JIG=17
            $ 192 "AMR_PosTarget≔5"
            global AMR_PosTarget=5
          else:
            $ 193 "ElseIf TASK.ID≟49"
            if (TASK.ID == 49):
              $ 194 "Task_info≔'Pick Containers'"
              global Task_info="Pick Containers"
              $ 195 "Parameters"
              $ 196 "ITM_ID≔1"
              global ITM_ID=1
              $ 197 "OBJ_Type≔6"
              global OBJ_Type=6
              $ 198 "JIG≔15"
              global JIG=15
              $ 199 "AMR_PosTarget≔3"
              global AMR_PosTarget=3
            else:
              $ 200 "ElseIf TASK.ID≟50"
              if (TASK.ID == 50):
                $ 201 "Task_info≔'Decap Containers'"
                global Task_info="Decap Containers"
                $ 202 "Parameters"
                $ 203 "ITM_ID≔1"
                global ITM_ID=1
                $ 204 "OBJ_Type≔6"
                global OBJ_Type=6
                $ 205 "JIG≔16"
                global JIG=16
                $ 206 "AMR_PosTarget≔5"
                global AMR_PosTarget=5
              else:
                $ 207 "ElseIf TASK.ID≟51"
                if (TASK.ID == 51):
                  $ 208 "Task_info≔'Detect Spatula and transfer powder'"
                  global Task_info="Detect Spatula and transfer powder"
                  $ 209 "Parameters"
                  $ 210 "ITM_ID≔1"
                  global ITM_ID=1
                  $ 211 "target_weight≔(UGO.read_input('00','Target_weight'))/1000"
                  global target_weight=(UGO.read_input("00","Target_weight"))/1000
                  $ 212 "OBJ_Type≔8"
                  global OBJ_Type=8
                  $ 213 "JIG≔16"
                  global JIG=16
                  $ 214 "AMR_PosTarget≔5"
                  global AMR_PosTarget=5
                else:
                  $ 215 "ElseIf TASK.ID≟52"
                  if (TASK.ID == 52):
                    $ 216 "Task_info≔'Pick Powder'"
                    global Task_info="Pick Powder"
                    $ 217 "Parameters"
                    $ 218 "ITM_ID≔1"
                    global ITM_ID=1
                    $ 220 "OBJ_Type≔6"
                    global OBJ_Type=6
                    $ 221 "JIG≔15"
                    global JIG=15
                    $ 222 "AMR_PosTarget≔3"
                    global AMR_PosTarget=3
                  else:
                    $ 223 "ElseIf TASK.ID≟53"
                    if (TASK.ID == 53):
                      $ 224 "Task_info≔'Decap Powder'"
                      global Task_info="Decap Powder"
                      $ 225 "Parameters"
                      $ 226 "ITM_ID≔1"
                      global ITM_ID=1
                      $ 227 "OBJ_Type≔6"
                      global OBJ_Type=6
                      $ 228 "JIG≔1"
                      global JIG=1
                      $ 229 "AMR_PosTarget≔5"
                      global AMR_PosTarget=5
                    else:
                      $ 230 "ElseIf TASK.ID≟54"
                      if (TASK.ID == 54):
                        $ 231 "Task_info≔'Empty and swap Powder container'"
                        global Task_info="Empty and swap Powder container"
                        $ 240 "Parameters"
                        $ 241 "ITM_ID≔1"
                        global ITM_ID=1
                        $ 243 "W_now≔(UGO.read_input('00','Container_weight'))/1000"
                        global W_now=(UGO.read_input("00","Container_weight"))/1000
                        $ 244 "Pow_name≔(UGO.read_input('00','Powder_name'))"
                        global Pow_name=(UGO.read_input("00","Powder_name"))
                        $ 247 "OBJ_Type≔6"
                        global OBJ_Type=6
                        $ 248 "JIG≔17"
                        global JIG=17
                        $ 249 "AMR_PosTarget≔5"
                        global AMR_PosTarget=5
                      else:
                        $ 250 "ElseIf TASK.ID≟55"
                        if (TASK.ID == 55):
                          $ 251 "Task_info≔'Place Powder'"
                          global Task_info="Place Powder"
                          $ 252 "Parameters"
                          $ 253 "ITM_ID≔1"
                          global ITM_ID=1
                          $ 254 "OBJ_Type≔6"
                          global OBJ_Type=6
                          $ 255 "JIG≔21"
                          global JIG=21
                          $ 256 "AMR_PosTarget≔5"
                          global AMR_PosTarget=5
                        else:
                          $ 257 "ElseIf TASK.ID≟56"
                          if (TASK.ID == 56):
                            $ 258 "Task_info≔'Dose Powder'"
                            global Task_info="Dose Powder"
                            $ 259 "Parameters"
                            $ 260 "ITM_ID≔1"
                            global ITM_ID=1
                            $ 261 "target_weight≔(UGO.read_input('00','Target_weight'))/1000"
                            global target_weight=(UGO.read_input("00","Target_weight"))/1000
                            $ 262 "W_now≔(UGO.read_input('00','Container_weight'))/1000"
                            global W_now=(UGO.read_input("00","Container_weight"))/1000
                            $ 263 "Pow_name≔(UGO.read_input('00','Powder_name'))"
                            global Pow_name=(UGO.read_input("00","Powder_name"))
                            $ 264 "OBJ_Type≔6"
                            global OBJ_Type=6
                            $ 265 "JIG≔17"
                            global JIG=17
                            $ 266 "AMR_PosTarget≔5"
                            global AMR_PosTarget=5
                          else:
                            $ 267 "ElseIf TASK.ID≟57"
                            if (TASK.ID == 57):
                              $ 268 "Task_info≔'Recipe Powder dosing'"
                              global Task_info="Recipe Powder dosing"
                              $ 269 "Parameters"
                              $ 270 "ITM_ID≔1"
                              global ITM_ID=1
                              $ 271 "Pow_A≔(UGO.read_input('00','PowderA'))"
                              global Pow_A=(UGO.read_input("00","PowderA"))
                              $ 272 "Pow_B≔(UGO.read_input('00','PowderB'))"
                              global Pow_B=(UGO.read_input("00","PowderB"))
                              $ 273 "Pow_C≔(UGO.read_input('00','PowderC'))"
                              global Pow_C=(UGO.read_input("00","PowderC"))
                              $ 274 "Total_weight≔(UGO.read_input('00','Total_weight'))/1000"
                              global Total_weight=(UGO.read_input("00","Total_weight"))/1000
                              $ 275 "Pow_A_percent≔(UGO.read_input('00','PowderA_percentage'))/100"
                              global Pow_A_percent=(UGO.read_input("00","PowderA_percentage"))/100
                              $ 276 "Pow_B_percent≔(UGO.read_input('00','PowderB_percentage'))/100"
                              global Pow_B_percent=(UGO.read_input("00","PowderB_percentage"))/100
                              $ 277 "Pow_C_percent≔(UGO.read_input('00','PowderC_percentage'))/100"
                              global Pow_C_percent=(UGO.read_input("00","PowderC_percentage"))/100
                              $ 278 "OBJ_Type≔6"
                              global OBJ_Type=6
                              $ 279 "JIG≔17"
                              global JIG=17
                              $ 280 "AMR_PosTarget≔5"
                              global AMR_PosTarget=5
                            else:
                              $ 281 "ElseIf TASK.ID≟58"
                              if (TASK.ID == 58):
                                $ 282 "Task_info≔'Pick Powder containers'"
                                global Task_info="Pick Powder containers"
                                $ 283 "Parameters"
                                $ 284 "ITM_ID≔1"
                                global ITM_ID=1
                                $ 285 "OBJ_Type≔6"
                                global OBJ_Type=6
                                $ 286 "JIG≔15"
                                global JIG=15
                                $ 287 "AMR_PosTarget≔3"
                                global AMR_PosTarget=3
                              else:
                                $ 288 "ElseIf TASK.ID≟59"
                                if (TASK.ID == 59):
                                  $ 289 "Task_info≔'Empty Powder container'"
                                  global Task_info="Empty Powder container"
                                  $ 290 "Parameters"
                                  $ 291 "ITM_ID≔1"
                                  global ITM_ID=1
                                  $ 293 "Pow_name≔(UGO.read_input('00','Powder_name'))"
                                  global Pow_name=(UGO.read_input("00","Powder_name"))
                                  $ 295 "target_weight≔(aa_weight_cont-empty_weight_g)*1000"
                                  global target_weight=(aa_weight_cont-empty_weight_g)*1000
                                  $ 296 "W_now≔target_weight"
                                  global W_now=target_weight
                                  $ 297 "send_picking_info(Pow_name,target_weight)"
                                  send_picking_info(Pow_name,target_weight)
                                  $ 298 "w_dosed_total≔0"
                                  global w_dosed_total=0
                                  $ 299 "OBJ_Type≔6"
                                  global OBJ_Type=6
                                  $ 300 "JIG≔17"
                                  global JIG=17
                                  $ 301 "AMR_PosTarget≔5"
                                  global AMR_PosTarget=5
                                else:
                                  $ 302 "ElseIf TASK.ID≟61"
                                  if (TASK.ID == 61):
                                    $ 303 "Task_info≔'Weigh, Place & Decap'"
                                    global Task_info="Weigh, Place & Decap"
                                    $ 304 "Parameters"
                                    $ 305 "ITM_ID≔1"
                                    global ITM_ID=1
                                    $ 306 "OBJ_Type≔6"
                                    global OBJ_Type=6
                                    $ 307 "JIG≔21"
                                    global JIG=21
                                    $ 308 "AMR_PosTarget≔5"
                                    global AMR_PosTarget=5
                                  else:
                                    $ 309 "ElseIf TASK.ID≟62"
                                    if (TASK.ID == 62):
                                      $ 310 "Task_info≔'Dose Powder'"
                                      global Task_info="Dose Powder"
                                      $ 311 "Parameters"
                                      $ 312 "ITM_ID≔1"
                                      global ITM_ID=1
                                      $ 314 "W_now≔aa_weight_cont"
                                      global W_now=aa_weight_cont
                                      $ 315 "Pow_name≔(UGO.read_input('00','Powder_name'))"
                                      global Pow_name=(UGO.read_input("00","Powder_name"))
                                      $ 316 "target_weight≔(UGO.read_input('00','Target_weight'))/1000"
                                      global target_weight=(UGO.read_input("00","Target_weight"))/1000
                                      $ 318 "params_init()"
                                      params_init()
                                      $ 319 "send_picking_info(Pow_name,target_weight)"
                                      send_picking_info(Pow_name,target_weight)
                                      $ 320 "OBJ_Type≔6"
                                      global OBJ_Type=6
                                      $ 321 "JIG≔17"
                                      global JIG=17
                                      $ 322 "AMR_PosTarget≔5"
                                      global AMR_PosTarget=5
                                    else:
                                      $ 323 "ElseIf TASK.ID≟63"
                                      if (TASK.ID == 63):
                                        $ 324 "Parameters"
                                        $ 325 "ITM_ID≔1"
                                        global ITM_ID=1
                                        $ 326 "OBJ_Type≔6"
                                        global OBJ_Type=6
                                        $ 327 "JIG≔21"
                                        global JIG=21
                                        $ 328 "AMR_PosTarget≔5"
                                        global AMR_PosTarget=5
                                      else:
                                        $ 329 "Else" "noBreak"
                                        $ 330 "set_error(ERROR_WRONG_ORDER)"
                                        set_error(ERROR_WRONG_ORDER)
                                      end
                                    end
                                  end
                                end
                              end
                            end
                          end
                        end
                      end
                    end
                  end
                end
              end
            end
          end
        end
      end
      $ 331 "test ugo"
      $ 332 "Wait: 0.2"
      sleep(0.2)
      $ 333 "ugo_update_outputs()"
      ugo_update_outputs()
      $ 334 "If starting() and AMR_Done"
      if (starting()  and  AMR_Done):
        $ 335 "log_message(Task_info, 'New Task: ')"
        log_message(Task_info, "New Task: ")
        $ 336 "log_message(to_str(TASK.ID), 'Task_ID: ')"
        log_message(to_str(TASK.ID), "Task_ID: ")
        $ 337 "do_transition(keep_rxry=OBJ_Picked)"
        do_transition(keep_rxry=OBJ_Picked)
        $ 338 "STATE≔6"
        global STATE=6
        $ 339 "ugo_update_outputs()"
        ugo_update_outputs()
      end
    elif (6 == switch_1):
      $ 340 "Case 6"
      $ 341 "Execute"
      $ 342 "STATE_Info≔'Execute'"
      global STATE_Info="Execute"
      $ 343 "If  not CMD_Hold and not CMD_Suspend"
      global thread_flag_343=0
      thread Thread_if_343():
        $ 344 "Switch PROCESS_Step"
        switch_2 = PROCESS_Step
        $ 345 "Case 0"
        if (0 == switch_2):
          $ 346 "PROCESS_Info≔'process control'"
          global PROCESS_Info="process control"
          $ 347 "log_process(PROCESS_Info)"
          log_process(PROCESS_Info)
          $ 348 "process control"
          $ 349 "If  not AMR_AtTarget"
          if (  not  AMR_AtTarget):
            $ 350 "PROCESS_Step≔1"
            global PROCESS_Step=1
          else:
            $ 351 "ElseIf (( not ITM_Prepared and  not WRK_Done) or (ITM_Prepared and WRK_Done))"
            if (((  not  ITM_Prepared  and    not  WRK_Done)  or  (ITM_Prepared  and  WRK_Done))):
              $ 352 "PROCESS_Step≔2"
              global PROCESS_Step=2
            else:
              $ 353 "ElseIf  not WRK_Done"
              if (  not  WRK_Done):
                $ 354 "PROCESS_Step≔3"
                global PROCESS_Step=3
              else:
                $ 355 "Else" "noBreak"
                $ 356 "task finished"
                $ 357 "PROCESS_Info≔''"
                global PROCESS_Info=""
                $ 358 "STATE≔7"
                global STATE=7
                $ 359 "ugo_update_outputs()"
                ugo_update_outputs()
              end
            end
          end
        elif (1 == switch_2):
          $ 360 "Case 1"
          $ 361 "navigate"
          $ 362 "'MOVING THE uML'"
          # 'MOVING THE uML'
          $ 363 "PROCESS_Info≔'move to target'"
          global PROCESS_Info="move to target"
          $ 364 "log_process(PROCESS_Info)"
          log_process(PROCESS_Info)
          $ 365 "If TASK.ID≟1"
          if (TASK.ID == 1):
            $ 366 "Action≔51"
            global Action=51
          else:
            $ 367 "Else" "noBreak"
            $ 368 "Action≔52"
            global Action=52
          end
          $ 369 "Call Sub_AMR_MiR_V3"
          Sub_AMR_MiR_V3()
          $ 370 "If AMR_Done"
          if (AMR_Done):
            $ 371 "PROCESS_Step≔0"
            global PROCESS_Step=0
          end
        elif (2 == switch_2):
          $ 372 "Case 2"
          $ 373 "prepare"
          $ 374 "'THINGS THAT HAVE TO BE DONE ONCE IN A SEQUENCE,WORKFLOW'"
          # 'THINGS THAT HAVE TO BE DONE ONCE IN A SEQUENCE,WORKFLOW'
          $ 375 "PROCESS_Info≔'prepare for work'"
          global PROCESS_Info="prepare for work"
          $ 376 "log_process(PROCESS_Info)"
          log_process(PROCESS_Info)
          $ 377 "If TASK.WORK.ITM_ID_Src>1"
          if (TASK.WORK.ITM_ID_Src>1):
            $ 378 "ITM_ID≔TASK.WORK.ITM_ID_Src"
            global ITM_ID=TASK.WORK.ITM_ID_Src
          else:
            $ 379 "ElseIf TASK.WORK.ITM_ID_Tgt>1"
            if (TASK.WORK.ITM_ID_Tgt>1):
              $ 380 "ITM_ID≔TASK.WORK.ITM_ID_Tgt"
              global ITM_ID=TASK.WORK.ITM_ID_Tgt
            end
          end
          $ 381 "If  not ARM_Referenced and (ITM_ID≠0)"
          if (  not  ARM_Referenced  and  (ITM_ID != 0)):
            $ 382 "STP≔1"
            global STP=1
          else:
            $ 383 "ElseIf ARM_Referenced or (ITM_ID≟0)"
            if (ARM_Referenced  or  (ITM_ID == 0)):
              $ 384 "STP≔2"
              global STP=2
            end
          end
          $ 385 "Switch STP"
          switch_3 = STP
          $ 386 "Case 1"
          if (1 == switch_3):
            $ 387 "reference"
            $ 388 "STP_Info≔'reference at target position'"
            global STP_Info="reference at target position"
            $ 389 "log_step(STP_Info)"
            log_step(STP_Info)
            $ 390 "If ITM_ID≟1"
            if (ITM_ID == 1):
              $ 391 "CAM_Done≔ True "
              global CAM_Done=  True
            else:
              $ 392 "Else" "noBreak"
              $ 393 "Action≔131"
              global Action=131
              $ 394 "Call Sub_Vision_V18"
              Sub_Vision_V18()
            end
            $ 396 "If CAM_Done and  not ERROR.FLAG"
            if (CAM_Done  and    not  ERROR.FLAG):
              $ 397 "log_step('ARM referenced')"
              log_step("ARM referenced")
              $ 398 "ARM_Referenced≔ True "
              global ARM_Referenced=  True
            end
          elif (2 == switch_3):
            $ 399 "Case 2"
            $ 400 "manipulate"
            $ 401 "STP_Info≔'manipulate item'"
            global STP_Info="manipulate item"
            $ 402 "log_step(STP_Info)"
            log_step(STP_Info)
            $ 403 "'In case pressing button is needed'"
            # 'In case pressing button is needed'
            $ 404 "If found_in_list(ITM_ID, ITM_ID_List)"
            if (found_in_list(ITM_ID, ITM_ID_List)):
              $ 405 "Switch ITM_ID"
              switch_4 = ITM_ID
              $ 406 "Case 0"
              if (0 == switch_4):
                $ 407 "ITM_Manipulated≔ not ITM_Manipulated"
                global ITM_Manipulated=  not  ITM_Manipulated
              elif (1 == switch_4):
                $ 408 "Case 1"
                $ 409 "ITM_Manipulated≔ not ITM_Manipulated"
                global ITM_Manipulated=  not  ITM_Manipulated
              elif (2 == switch_4):
                $ 410 "Case 2"
              else:
                $ 420 "Default Case"
                $ 421 "ITM_Manipulated≔ not ITM_Manipulated"
                global ITM_Manipulated=  not  ITM_Manipulated
              end
            end
          end
          $ 422 "ITM_Prepared≔(ITM_Manipulated or  not found_in_list(ITM_ID, ITM_ID_List)) and (ARM_Referenced or ITM_ID≟0) and  not WRK_Done"
          global ITM_Prepared=(ITM_Manipulated  or    not  found_in_list(ITM_ID, ITM_ID_List))  and  (ARM_Referenced  or  ITM_ID == 0)  and    not  WRK_Done
          $ 423 "STP≔0"
          global STP=0
          $ 424 "STP_Info≔''"
          global STP_Info=""
          $ 425 "PROCESS_Step≔0"
          global PROCESS_Step=0
        elif (3 == switch_2):
          $ 426 "Case 3"
          $ 427 "work"
          $ 428 "'ADD EVERY MACHINE, OBJECT, STATION TO WORK ON'"
          # 'ADD EVERY MACHINE, OBJECT, STATION TO WORK ON'
          $ 429 "Switch ITM_ID"
          switch_3 = ITM_ID
          $ 430 "Case 1"
          if (1 == switch_3):
            $ 431 "uLM"
            $ 432 "If TASK.ID≟12"
            if (TASK.ID == 12):
              $ 433 "fill racks"
              $ 434 "Action≔151"
              global Action=151
              $ 435 "Call Sub_Vision_V18"
              Sub_Vision_V18()
              $ 436 "If  not ERROR.FLAG"
              if (  not  ERROR.FLAG):
                $ 437 "Actions for the task"
                $ 438 "Action≔1"
                global Action=1
                $ 439 "JIG≔2"
                global JIG=2
                $ 440 "JIG_Slot≔CAM_Result[0]"
                global JIG_Slot=CAM_Result[0]
                $ 441 "OBJ_Nbr≔CAM_Result[0]"
                global OBJ_Nbr=CAM_Result[0]
                $ 442 "OBJ_Type≔2"
                global OBJ_Type=2
                $ 443 "Call Sub_Action_V4"
                Sub_Action_V4()
                $ 444 "If OBJ_Picked"
                if (OBJ_Picked):
                  $ 445 "CAM_Result.remove(0)"
                  CAM_Result.remove(0)
                  $ 446 "PRC_TubCounter≔PRC_TubCounter+1"
                  global PRC_TubCounter=PRC_TubCounter+1
                  $ 447 "If PRC_TubCounter%4≟0"
                  if (PRC_TubCounter%4 == 0):
                    $ 448 "JIG_Slot≔4"
                    global JIG_Slot=4
                  else:
                    $ 449 "Else" "noBreak"
                    $ 450 "JIG_Slot≔PRC_TubCounter%4"
                    global JIG_Slot=PRC_TubCounter%4
                  end
                  $ 451 "OBJ_Nbr≔ceil(PRC_TubCounter/4)"
                  global OBJ_Nbr=ceil(PRC_TubCounter/4)
                  $ 452 "Action≔2"
                  global Action=2
                  $ 453 "JIG≔4"
                  global JIG=4
                  $ 454 "Call Sub_Action_V4"
                  Sub_Action_V4()
                  $ 455 "Action≔151"
                  global Action=151
                  $ 456 "Call Sub_Vision_V18"
                  Sub_Vision_V18()
                end
              end
              $ 457 "If (CAM_Captures≥CAM_PRM_Retries) or (PRC_TubCounter≥32)"
              if ((CAM_Captures >= CAM_PRM_Retries)  or  (PRC_TubCounter >= 32)):
                $ 458 "PROCESS_Step≔0"
                global PROCESS_Step=0
                $ 459 "WRK_Done≔ True "
                global WRK_Done=  True
              end
            else:
              $ 460 "ElseIf TASK.ID≟13"
              if (TASK.ID == 13):
                $ 461 "Dose Powder"
                $ 462 "Action≔131"
                global Action=131
                $ 463 "Call Sub_Vision_V18"
                Sub_Vision_V18()
                $ 464 "Action≔34"
                global Action=34
                $ 465 "Call Sub_Action_V4"
                Sub_Action_V4()
                $ 466 "PROCESS_Step≔0"
                global PROCESS_Step=0
                $ 467 "WRK_Done≔ True "
                global WRK_Done=  True
              else:
                $ 468 "ElseIf TASK.ID≟49"
                if (TASK.ID == 49):
                  $ 469 "Pick Powder container"
                  $ 470 "Action≔131"
                  global Action=131
                  $ 471 "Call Sub_Vision_V18"
                  Sub_Vision_V18()
                  $ 472 "Action≔35"
                  global Action=35
                  $ 473 "Call Sub_Action_V4"
                  Sub_Action_V4()
                  $ 474 "PROCESS_Step≔0"
                  global PROCESS_Step=0
                  $ 475 "WRK_Done≔ True "
                  global WRK_Done=  True
                else:
                  $ 476 "ElseIf TASK.ID≟50"
                  if (TASK.ID == 50):
                    $ 477 "Decap containers"
                    $ 478 "Action≔36"
                    global Action=36
                    $ 479 "Call Sub_Action_V4"
                    Sub_Action_V4()
                    $ 480 "PROCESS_Step≔0"
                    global PROCESS_Step=0
                    $ 481 "WRK_Done≔ True "
                    global WRK_Done=  True
                  else:
                    $ 482 "ElseIf TASK.ID≟51"
                    if (TASK.ID == 51):
                      $ 483 "Detect Spatula and transfer powder"
                      $ 484 "Action≔131"
                      global Action=131
                      $ 485 "Call Sub_Vision_V18"
                      Sub_Vision_V18()
                      $ 486 "Action≔37"
                      global Action=37
                      $ 487 "Call Sub_Action_V4"
                      Sub_Action_V4()
                      $ 488 "PROCESS_Step≔0"
                      global PROCESS_Step=0
                      $ 489 "WRK_Done≔ True "
                      global WRK_Done=  True
                    else:
                      $ 490 "ElseIf TASK.ID≟52"
                      if (TASK.ID == 52):
                        $ 491 "Pick Powder container"
                        $ 492 "Action≔131"
                        global Action=131
                        $ 493 "Call Sub_Vision_V18"
                        Sub_Vision_V18()
                        $ 494 "Action≔39"
                        global Action=39
                        $ 495 "Call Sub_Action_V4"
                        Sub_Action_V4()
                        $ 496 "PROCESS_Step≔0"
                        global PROCESS_Step=0
                        $ 497 "WRK_Done≔ True "
                        global WRK_Done=  True
                      else:
                        $ 498 "ElseIf TASK.ID≟53"
                        if (TASK.ID == 53):
                          $ 499 "Decap containerA"
                          $ 500 "Action≔40"
                          global Action=40
                          $ 501 "Call Sub_Action_V4"
                          Sub_Action_V4()
                          $ 502 "PROCESS_Step≔0"
                          global PROCESS_Step=0
                          $ 503 "WRK_Done≔ True "
                          global WRK_Done=  True
                        else:
                          $ 504 "ElseIf TASK.ID≟55"
                          if (TASK.ID == 55):
                            $ 505 "Place Powder"
                            $ 506 "Action≔131"
                            global Action=131
                            $ 507 "Call Sub_Vision_V18"
                            Sub_Vision_V18()
                            $ 508 "Action≔41"
                            global Action=41
                            $ 509 "Call Sub_Action_V4"
                            Sub_Action_V4()
                            $ 510 "PROCESS_Step≔0"
                            global PROCESS_Step=0
                            $ 511 "WRK_Done≔ True "
                            global WRK_Done=  True
                          else:
                            $ 512 "ElseIf TASK.ID≟54"
                            if (TASK.ID == 54):
                              $ 513 "Empty and swap container"
                              $ 514 "Action≔131"
                              global Action=131
                              $ 515 "Call Sub_Vision_V18"
                              Sub_Vision_V18()
                              $ 516 "Action≔42"
                              global Action=42
                              $ 517 "Call Sub_Action_V4"
                              Sub_Action_V4()
                              $ 518 "PROCESS_Step≔0"
                              global PROCESS_Step=0
                              $ 519 "WRK_Done≔ True "
                              global WRK_Done=  True
                            else:
                              $ 520 "ElseIf TASK.ID≟56"
                              if (TASK.ID == 56):
                                $ 521 "Dispense Powder"
                                $ 522 "Action≔131"
                                global Action=131
                                $ 523 "Call Sub_Vision_V18"
                                Sub_Vision_V18()
                                $ 524 "Action≔43"
                                global Action=43
                                $ 525 "Call Sub_Action_V4"
                                Sub_Action_V4()
                                $ 526 "PROCESS_Step≔0"
                                global PROCESS_Step=0
                                $ 527 "WRK_Done≔ True "
                                global WRK_Done=  True
                              else:
                                $ 528 "ElseIf TASK.ID≟57"
                                if (TASK.ID == 57):
                                  $ 529 "Recipe Dosing"
                                  $ 530 "Action≔48"
                                  global Action=48
                                  $ 531 "Call Sub_Action_V4"
                                  Sub_Action_V4()
                                  $ 548 "PROCESS_Step≔0"
                                  global PROCESS_Step=0
                                  $ 549 "WRK_Done≔ True "
                                  global WRK_Done=  True
                                else:
                                  $ 550 "ElseIf TASK.ID≟58"
                                  if (TASK.ID == 58):
                                    $ 551 "Pick Powder containers"
                                    $ 552 "Num_cont_picked≔0"
                                    global Num_cont_picked=0
                                    $ 553 "powder_position≔'Position1'"
                                    global powder_position="Position1"
                                    $ 554 "Loop Num_cont_picked<3"
                                    while (Num_cont_picked<3):
                                      $ 555 "Action≔131"
                                      global Action=131
                                      $ 556 "Call Sub_Vision_V18"
                                      Sub_Vision_V18()
                                      $ 557 "Action≔47"
                                      global Action=47
                                      $ 558 "Call Sub_Action_V4"
                                      Sub_Action_V4()
                                    end
                                    $ 559 "PROCESS_Step≔0"
                                    global PROCESS_Step=0
                                    $ 560 "WRK_Done≔ True "
                                    global WRK_Done=  True
                                  else:
                                    $ 561 "ElseIf TASK.ID≟59"
                                    if (TASK.ID == 59):
                                      $ 562 "Empty powder container"
                                      $ 563 "Action≔131"
                                      global Action=131
                                      $ 564 "Call Sub_Vision_V18"
                                      Sub_Vision_V18()
                                      $ 565 "Action≔50"
                                      global Action=50
                                      $ 566 "Call Sub_Action_V4"
                                      Sub_Action_V4()
                                      $ 567 "PROCESS_Step≔0"
                                      global PROCESS_Step=0
                                      $ 568 "WRK_Done≔ True "
                                      global WRK_Done=  True
                                    else:
                                      $ 569 "ElseIf TASK.ID≟61"
                                      if (TASK.ID == 61):
                                        $ 570 "Place Powder"
                                        $ 571 "Action≔131"
                                        global Action=131
                                        $ 572 "Call Sub_Vision_V18"
                                        Sub_Vision_V18()
                                        $ 573 "Action≔51"
                                        global Action=51
                                        $ 574 "Call Sub_Action_V4"
                                        Sub_Action_V4()
                                        $ 575 "PROCESS_Step≔0"
                                        global PROCESS_Step=0
                                        $ 576 "WRK_Done≔ True "
                                        global WRK_Done=  True
                                      else:
                                        $ 577 "ElseIf TASK.ID≟62"
                                        if (TASK.ID == 62):
                                          $ 578 "Dose Powder"
                                          $ 579 "Action≔131"
                                          global Action=131
                                          $ 580 "Call Sub_Vision_V18"
                                          Sub_Vision_V18()
                                          $ 581 "Action≔52"
                                          global Action=52
                                          $ 582 "Call Sub_Action_V4"
                                          Sub_Action_V4()
                                          $ 583 "PROCESS_Step≔0"
                                          global PROCESS_Step=0
                                          $ 584 "WRK_Done≔ True "
                                          global WRK_Done=  True
                                        else:
                                          $ 585 "ElseIf TASK.ID≟63"
                                          if (TASK.ID == 63):
                                            $ 586 "Swabbing"
                                            $ 587 "Action≔131"
                                            global Action=131
                                            $ 588 "Call Sub_Vision_V18"
                                            Sub_Vision_V18()
                                            $ 589 "Action≔53"
                                            global Action=53
                                            $ 590 "Call Sub_Action_V4"
                                            Sub_Action_V4()
                                            $ 591 "PROCESS_Step≔0"
                                            global PROCESS_Step=0
                                            $ 592 "WRK_Done≔ True "
                                            global WRK_Done=  True
                                          end
                                        end
                                      end
                                    end
                                  end
                                end
                              end
                            end
                          end
                        end
                      end
                    end
                  end
                end
              end
            end
          elif (2 == switch_3):
            $ 593 "Case 2"
          elif (5 == switch_3):
            $ 635 "Case 5"
          elif (20 == switch_3):
            $ 643 "Case 20"
          elif (43 == switch_3):
            $ 705 "Case 43"
          else:
            $ 713 "Default Case"
            $ 714 "WRK_Done≔ True "
            global WRK_Done=  True
            $ 715 "PROCESS_Step≔0"
            global PROCESS_Step=0
          end
        end
        thread_flag_343 = 1
      end
      if (  not  CMD_Hold and not CMD_Suspend):
        global thread_handler_343=run Thread_if_343()
        while (thread_flag_343 == 0):
          if not(  not  CMD_Hold and not CMD_Suspend):
            kill thread_handler_343
            thread_flag_343 = 2
          else:
            sync()
          end
        end
      else:
        thread_flag_343 = 2
      end
      $ 716 "If CMD_Hold"
      if (CMD_Hold):
        $ 717 "STATE≔9"
        global STATE=9
        $ 718 "ugo_update_outputs()"
        ugo_update_outputs()
      else:
        $ 719 "ElseIf CMD_Suspend"
        if (CMD_Suspend):
          $ 720 "STATE≔12"
          global STATE=12
          $ 721 "ugo_update_outputs()"
          ugo_update_outputs()
        end
      end
    elif (7 == switch_1):
      $ 722 "Case 7"
      $ 723 "Completing"
      $ 724 "STATE_Info≔'Completing'"
      global STATE_Info="Completing"
      $ 725 "'ADD COMMANDS FOR COMPLETING THE PROCESS'"
      # 'ADD COMMANDS FOR COMPLETING THE PROCESS'
      $ 726 "do_transition(keep_rxry=OBJ_Picked)"
      do_transition(keep_rxry=OBJ_Picked)
      $ 727 "Call Sub_AMR_MiR_V3"
      Sub_AMR_MiR_V3()
      $ 728 "If completing() and AMR_Done"
      if (completing()  and  AMR_Done):
        $ 729 "STATE≔8"
        global STATE=8
        $ 730 "ugo_update_outputs()"
        ugo_update_outputs()
      end
    elif (8 == switch_1):
      $ 731 "Case 8"
      $ 732 "Complete"
      $ 733 "STATE_Info≔'Complete'"
      global STATE_Info="Complete"
      $ 734 "If CMD_Reset"
      if (CMD_Reset):
        $ 735 "STATE≔3"
        global STATE=3
        $ 736 "ugo_update_outputs()"
        ugo_update_outputs()
      end
    elif (9 == switch_1):
      $ 737 "Case 9"
      $ 738 "Holding"
      $ 739 "STATE_Info≔'Holding'"
      global STATE_Info="Holding"
      $ 740 "stopl(0.5)"
      stopl(0.5)
      $ 741 "Call Sub_AMR_MiR_V3"
      Sub_AMR_MiR_V3()
      $ 742 "If holding() and AMR_Done"
      if (holding()  and  AMR_Done):
        $ 743 "STATE≔10"
        global STATE=10
        $ 744 "ugo_update_outputs()"
        ugo_update_outputs()
      end
    elif (10 == switch_1):
      $ 745 "Case 10"
      $ 746 "Held"
      $ 747 "STATE_Info≔'Held'"
      global STATE_Info="Held"
      $ 748 "If CMD_Unhold"
      if (CMD_Unhold):
        $ 749 "end_freedrive_mode()"
        end_freedrive_mode()
        $ 750 "STATE≔11"
        global STATE=11
        $ 751 "ugo_update_outputs()"
        ugo_update_outputs()
      else:
        $ 752 "ElseIf FNC_Freedrive"
        if (FNC_Freedrive):
          $ 753 "freedrive_mode()"
          freedrive_mode()
        else:
          $ 754 "Else" "noBreak"
          $ 755 "end_freedrive_mode()"
          end_freedrive_mode()
        end
      end
    elif (11 == switch_1):
      $ 756 "Case 11"
      $ 757 "Unholding"
      $ 758 "STATE_Info≔'Unholding'"
      global STATE_Info="Unholding"
      $ 759 "Clearing"
      $ 760 "Switch ERROR.ID"
      switch_2 = ERROR.ID
      $ 761 "Case 1002"
      if (1002 == switch_2):
        $ 762 "AMR_AtTarget≔ False "
        global AMR_AtTarget=  False
        $ 763 "ARM_Referenced≔ False "
        global ARM_Referenced=  False
        $ 764 "ITM_Prepared≔ False "
        global ITM_Prepared=  False
        $ 765 "PROCESS_Step≔1"
        global PROCESS_Step=1
      elif (2007 == switch_2):
        $ 766 "Case 2007"
        $ 767 "PROCESS_Step≔1"
        global PROCESS_Step=1
      end
      $ 768 "reset_error()"
      reset_error()
      $ 769 "reset_warning()"
      reset_warning()
      $ 770 "OBJ_Picked≔gripper_has_object()"
      global OBJ_Picked=gripper_has_object()
      $ 771 "Call Sub_AMR_MiR_V3"
      Sub_AMR_MiR_V3()
      $ 772 "If unholding() and AMR_Done"
      if (unholding()  and  AMR_Done):
        $ 773 "STATE≔6"
        global STATE=6
        $ 774 "ugo_update_outputs()"
        ugo_update_outputs()
      end
    elif (12 == switch_1):
      $ 775 "Case 12"
      $ 776 "Suspending"
      $ 777 "STATE_Info≔'Suspending'"
      global STATE_Info="Suspending"
      $ 778 "PROCESS_Info≔str_cat(PROCESS_Info, ' suspended')"
      global PROCESS_Info=str_cat(PROCESS_Info, " suspended")
      $ 779 "If suspending()"
      if (suspending()):
        $ 780 "STATE≔13"
        global STATE=13
        $ 781 "ugo_update_outputs()"
        ugo_update_outputs()
      end
    elif (13 == switch_1):
      $ 782 "Case 13"
      $ 783 "Suspended"
      $ 784 "STATE_Info≔'Suspended'"
      global STATE_Info="Suspended"
      $ 785 "Call Sub_AMR_MiR_V3"
      Sub_AMR_MiR_V3()
      $ 786 "If CMD_Unsuspend"
      if (CMD_Unsuspend):
        $ 787 "STATE≔14"
        global STATE=14
        $ 788 "ugo_update_outputs()"
        ugo_update_outputs()
      end
    elif (14 == switch_1):
      $ 789 "Case 14"
      $ 790 "Unsuspending"
      $ 791 "STATE_Info≔'Unsuspending'"
      global STATE_Info="Unsuspending"
      $ 792 "PROCESS_Step≔0"
      global PROCESS_Step=0
      $ 793 "If unsuspending()"
      if (unsuspending()):
        $ 794 "STATE≔6"
        global STATE=6
        $ 795 "ugo_update_outputs()"
        ugo_update_outputs()
      end
    elif (15 == switch_1):
      $ 796 "Case 15"
      $ 797 "Aborting"
      $ 798 "STATE_Info≔'Aborting'"
      global STATE_Info="Aborting"
      $ 799 "If aborting()"
      if (aborting()):
        $ 800 "STATE≔16"
        global STATE=16
        $ 801 "ugo_update_outputs()"
        ugo_update_outputs()
      end
    elif (16 == switch_1):
      $ 802 "Case 16"
      $ 803 "Aborted"
      $ 804 "STATE_Info≔'Aborted'"
      global STATE_Info="Aborted"
      $ 805 "If CMD_Clear"
      if (CMD_Clear):
        $ 806 "STATE≔17"
        global STATE=17
        $ 807 "ugo_update_outputs()"
        ugo_update_outputs()
      end
    elif (17 == switch_1):
      $ 808 "Case 17"
      $ 809 "Clearing"
      $ 810 "STATE_Info≔'Clearing'"
      global STATE_Info="Clearing"
      $ 811 "Clearing"
      $ 812 "reset_warning()"
      reset_warning()
      $ 813 "reset_error()"
      reset_error()
      $ 814 "If clearing()"
      if (clearing()):
        $ 815 "STATE≔2"
        global STATE=2
        $ 816 "ugo_update_outputs()"
        ugo_update_outputs()
      end
    end
    $ 817 "log_state(STATE_Info)"
    log_state(STATE_Info)
    $ 818 "log_warning(WARNING.MSG)"
    log_warning(WARNING.MSG)
    $ 819 "log_error(ERROR.MSG)"
    log_error(ERROR.MSG)
    $ 820 "Times"
    $ 821 "Switch STATE"
    switch_1 = STATE
    $ 822 "Case 1"
    if (1 == switch_1):
      $ 823 "TM_St_Stopping≔get_time(STATE_Times[STATE-1])"
      global TM_St_Stopping=get_time(STATE_Times[STATE-1])
    elif (2 == switch_1):
      $ 824 "Case 2"
      $ 825 "TM_St_Stopped≔get_time(STATE_Times[STATE-1])"
      global TM_St_Stopped=get_time(STATE_Times[STATE-1])
    elif (3 == switch_1):
      $ 826 "Case 3"
      $ 827 "TM_St_Resetting≔get_time(STATE_Times[STATE-1])"
      global TM_St_Resetting=get_time(STATE_Times[STATE-1])
    elif (4 == switch_1):
      $ 828 "Case 4"
      $ 829 "TM_St_Idle≔get_time(STATE_Times[STATE-1])"
      global TM_St_Idle=get_time(STATE_Times[STATE-1])
    elif (5 == switch_1):
      $ 830 "Case 5"
      $ 831 "TM_St_Starting≔get_time(STATE_Times[STATE-1])"
      global TM_St_Starting=get_time(STATE_Times[STATE-1])
    elif (6 == switch_1):
      $ 832 "Case 6"
      $ 833 "TM_St_Execute≔get_time(STATE_Times[STATE-1])"
      global TM_St_Execute=get_time(STATE_Times[STATE-1])
    elif (7 == switch_1):
      $ 834 "Case 7"
      $ 835 "TM_St_Completin≔get_time(STATE_Times[STATE-1])"
      global TM_St_Completin=get_time(STATE_Times[STATE-1])
    elif (8 == switch_1):
      $ 836 "Case 8"
      $ 837 "TM_St_Complete≔get_time(STATE_Times[STATE-1])"
      global TM_St_Complete=get_time(STATE_Times[STATE-1])
    elif (9 == switch_1):
      $ 838 "Case 9"
      $ 839 "TM_St_Holding≔get_time(STATE_Times[STATE-1])"
      global TM_St_Holding=get_time(STATE_Times[STATE-1])
    elif (10 == switch_1):
      $ 840 "Case 10"
      $ 841 "TM_St_Held≔get_time(STATE_Times[STATE-1])"
      global TM_St_Held=get_time(STATE_Times[STATE-1])
    elif (11 == switch_1):
      $ 842 "Case 11"
      $ 843 "TM_St_Unholding≔get_time(STATE_Times[STATE-1])"
      global TM_St_Unholding=get_time(STATE_Times[STATE-1])
    elif (12 == switch_1):
      $ 844 "Case 12"
      $ 845 "TM_St_Suspendin≔get_time(STATE_Times[STATE-1])"
      global TM_St_Suspendin=get_time(STATE_Times[STATE-1])
    elif (13 == switch_1):
      $ 846 "Case 13"
      $ 847 "TM_St_Suspended≔get_time(STATE_Times[STATE-1])"
      global TM_St_Suspended=get_time(STATE_Times[STATE-1])
    elif (14 == switch_1):
      $ 848 "Case 14"
      $ 849 "TM_St_Unsuspend≔get_time(STATE_Times[STATE-1])"
      global TM_St_Unsuspend=get_time(STATE_Times[STATE-1])
    elif (15 == switch_1):
      $ 850 "Case 15"
      $ 851 "TM_St_Aborting≔get_time(STATE_Times[STATE-1])"
      global TM_St_Aborting=get_time(STATE_Times[STATE-1])
    elif (16 == switch_1):
      $ 852 "Case 16"
      $ 853 "TM_St_Aborted≔get_time(STATE_Times[STATE-1])"
      global TM_St_Aborted=get_time(STATE_Times[STATE-1])
    elif (17 == switch_1):
      $ 854 "Case 17"
      $ 855 "TM_St_Clearing≔get_time(STATE_Times[STATE-1])"
      global TM_St_Clearing=get_time(STATE_Times[STATE-1])
    end
    $ 857 "Wait: 0.1"
    sleep(0.1)
  end
end
